(* IEC 61131-3 sources: daoli-st-library/_tmp_r79, 4 files *)

(* ---- probe_idioms3.st ---- *)
FUNCTION FC_DL_ProbeF : DINT
VAR_INPUT
    nMonth : DINT;                   // 月 / month
    bLeap : BOOL;                    // 闰年 / leap year
END_VAR
VAR
    nDays : DINT;                    // 天数 / days
    i : DINT;                        // 索引 / index
    nSum : DINT;                     // 和 / sum
    nCnt : DINT;                     // 计数 / count
END_VAR
nDays := 0;
CASE nMonth OF
    1, 3, 5, 7, 8, 10, 12:
        nDays := 31;
    4, 6, 9, 11:
        nDays := 30;
    2:
        IF bLeap THEN
            nDays := 29;
        ELSE
            nDays := 28;
        END_IF
ELSE
    nDays := 0;
END_CASE
nSum := 0;
nCnt := 0;
FOR i := 1 TO 10 DO
    nCnt := nCnt + 1;
    IF nCnt > 5 THEN
        EXIT;
    END_IF
    nSum := nSum + i;
END_FOR
WHILE (nSum > 0) AND (nCnt < 30) DO
    nSum := nSum - 1;
    nCnt := nCnt + 1;
END_WHILE
IF (nDays = 0) THEN
    FC_DL_ProbeF := nSum;
    RETURN;
END_IF
FC_DL_ProbeF := nDays + nCnt;
END_FUNCTION

(* ---- probe_idioms4.st ---- *)
FUNCTION FC_DL_ProbeG : DINT
VAR_INPUT
    nA : DINT;                       // 输入 / input
END_VAR
VAR
    nB : DINT;                       // 中间量 / intermediate
    nC : DINT;                       // 中间量二 / second intermediate
END_VAR
nB := 1; nC := 2;
IF nA > 0 THEN
    nB := 3; nC := 4;
ELSE
    nB := 5; nC := 6;
END_IF
FC_DL_ProbeG := nB + nC;
END_FUNCTION

(* ---- probe_idioms.st ---- *)
FUNCTION FC_DL_ProbeA : LREAL
VAR_INPUT
    aPtsX : ARRAY[1..10] OF LREAL;   // 探针 X 数组 / probe X array
    aPtsY : ARRAY[1..10] OF LREAL;   // 探针 Y 数组 / probe Y array
    nCnt : INT;                      // 点数 / point count
END_VAR
VAR_OUTPUT
    eErr : UDINT;                    // 错误码 / error id
    bError : BOOL;                   // 故障标志 / fault flag
    bValid : BOOL;                   // 有效标志 / valid flag
END_VAR
VAR
    fSum : LREAL;                    // 累计 / accumulator
    fDx : LREAL;                     // 差值 / delta
    i : INT;                         // 索引 / index
    nB : UDINT;                      // 探针无符号 / probe unsigned
    nC : UDINT;                      // 探针无符号二 / probe unsigned two
    nD : UDINT;                      // 探针无符号三 / probe unsigned three
END_VAR
VAR CONSTANT
    DL_EPS : LREAL := 1.0E-9;        // 容差 / epsilon
    DL_MAX : UDINT := 16#FFFF_FFFF;  // 上限 / upper bound
END_VAR
fSum := 0.0;
eErr := 0;
bError := FALSE;
bValid := TRUE;
FOR i := 1 TO 10 DO
    fDx := aPtsX[i] - aPtsY[i];
    fSum := fSum + SQRT(fDx * fDx + DL_EPS);
END_FOR
nB := 123456;
nC := nB / 10;
nD := nB MOD 10;
IF nD > DL_MAX THEN
    bError := TRUE;
END_IF
IF EXPT(2.0, 3.0) > 7.0 THEN
    fSum := fSum + ATAN(1.0);
END_IF
FC_DL_ProbeA := fSum + LREAL_TO_REAL(fSum);
END_FUNCTION

FUNCTION FC_DL_ProbeB : UDINT
VAR_INPUT
    nVal : UDINT;                    // 探针输入 / probe input
END_VAR
VAR_OUTPUT
    eErr : UDINT;                    // 错误码 / error id
    bError : BOOL;                   // 故障标志 / fault flag
    bOverflow : BOOL;                // 溢出标志 / overflow flag
END_VAR
VAR
    nRoot : UDINT;                   // 试根 / trial root
    nIter : UDINT;                   // 迭代计数 / iteration counter
    fTmp : LREAL;                    // 探针实数 / probe real
END_VAR
nRoot := nVal;
nIter := 0;
WHILE (nIter < 64) AND (nRoot > 1) DO
    nRoot := nRoot / 2;
    nIter := nIter + 1;
END_WHILE
fTmp := TRUNC(LREAL_TO_REAL(1.5));
FC_DL_ProbeB := nRoot + LREAL_TO_UDINT(fTmp);
END_FUNCTION

FUNCTION_BLOCK FB_DL_ProbeC
VAR_INPUT
    bEnable : BOOL;                  // 使能 / enable
    bReset : BOOL;                   // 复位上升沿 / reset rising edge
    fSample : LREAL;                 // 样本 / sample
END_VAR
VAR_OUTPUT
    fMean : LREAL;                   // 均值 / mean
    nCount : UDINT;                  // 计数 / count
END_VAR
VAR
    rtReset : R_TRIG;                // 复位沿 / reset edge
    nStep : INT;                     // 内部状态 / internal state
    fSum : LREAL;                    // 累计 / accumulator
END_VAR
VAR CONSTANT
    DL_NAN_GUARD : LREAL := 1.0E308; // 有限上限 / finite ceiling
END_VAR
rtReset(CLK := bReset);
IF rtReset.Q THEN
    fSum := 0.0;
    nCount := 0;
    nStep := 0;
END_IF
CASE nStep OF
    0:
        IF bEnable THEN
            nStep := 10;
        END_IF
    10:
        IF NOT ((fSample <> fSample) OR (ABS(fSample) > DL_NAN_GUARD)) THEN
            fSum := fSum + fSample;
            nCount := nCount + 1;
            IF nCount > 0 THEN
                fMean := fSum / UDINT_TO_LREAL(nCount);
            END_IF
        END_IF
ELSE
    nStep := 0;
END_CASE
END_FUNCTION_BLOCK

(* ---- probe_idioms2.st ---- *)
TYPE E_DL_ProbeState :
(
    eIdle := 0,          // 空闲 / idle
    eRun := 1            // 运行 / run
);
END_TYPE

FUNCTION FC_DL_ProbeD : UDINT
VAR_INPUT
    aData : ARRAY[1..16] OF BYTE;    // 字节块 / byte block
    nLen : INT;                      // 长度 / length
END_VAR
VAR_OUTPUT
    eErr : UDINT;                    // 错误码 / error id
    bError : BOOL;                   // 故障标志 / fault flag
END_VAR
VAR
    nSum1 : UDINT;                   // 和 1 / sum one
    nSum2 : UDINT;                   // 和 2 / sum two
    nByte : UDINT;                   // 字节值 / byte value
    nWord : UDINT;                   // 字值 / word value
    nLo : UDINT;                     // 低字节 / low byte
    nHi : UDINT;                     // 高字节 / high byte
    bTmp : BYTE;                     // 字节中间量 / byte intermediate
    i : INT;                         // 索引 / index
    nUse : INT;                      // 有效长度 / effective length
END_VAR
VAR CONSTANT
    DL_MOD : UDINT := 255;           // 模数 / modulus
    DL_SHIFT : UDINT := 8;           // 移位量 / shift amount
END_VAR
eErr := 0;
bError := FALSE;
nSum1 := 0;
nSum2 := 0;
nUse := nLen;
IF nUse < 0 THEN
    nUse := 0;
ELSIF nUse > 16 THEN
    nUse := 16;
END_IF
FOR i := 1 TO nUse DO
    nByte := BYTE_TO_UDINT(aData[i]);
    nSum1 := (nSum1 + nByte) MOD DL_MOD;
    nSum2 := (nSum2 + nSum1) MOD DL_MOD;
END_FOR
nLo := BYTE_TO_UDINT(aData[1]);
nHi := BYTE_TO_UDINT(aData[2]);
nWord := nLo + nHi * 256;
bTmp := UDINT_TO_BYTE(nWord MOD DL_MOD);
FC_DL_ProbeD := (nSum2 * 256 + nSum1) + BYTE_TO_UDINT(bTmp) + nWord * 0;
END_FUNCTION

FUNCTION_BLOCK FB_DL_ProbeE
VAR_INPUT
    bEnable : BOOL;                  // 使能 / enable
END_VAR
VAR_OUTPUT
    eState : E_DL_ProbeState;        // 状态 / state
END_VAR
VAR
    nIdx : UDINT;                    // 计数 / counter
    nA : UDINT;                      // 无符号一 / unsigned one
    nB : UDINT;                      // 无符号二 / unsigned two
    nQ : DINT;                       // 有符号商 / signed quotient
    nR : DINT;                       // 有符号余 / signed remainder
END_VAR
VAR CONSTANT
    DL_DINT_MIN_P : DINT := -2147483648;  // 下界 / lower bound
    DL_DINT_MAX_P : DINT := 2147483647;   // 上界 / upper bound
END_VAR
eState := eIdle;
nA := 16#FFFF_FFFF;
nB := 0;
IF bEnable THEN
    eState := eRun;
    nB := nA / 2;
    nIdx := nA - nB;
    IF (nIdx > 1000) AND (nIdx < 16#FFFF_FFFF) THEN
        nQ := UDINT_TO_DINT(nIdx);
        nR := nQ MOD 7;
    END_IF
END_IF
IF (nQ = DL_DINT_MIN_P) OR (nR = DL_DINT_MAX_P) THEN
    eState := eIdle;
END_IF
IF eState = eRun THEN
    nIdx := nIdx + 1;
END_IF
END_FUNCTION_BLOCK
